DATA_BLOCK "GDB_PressDemoHardwareDriver"
{ S7_Optimized_Access := 'TRUE' }
VERSION : 0.1
NON_RETAIN
"FB_PressDemoHardwareDriver"
BEGIN
END_DATA_BLOCK
